TYPE ST_MotorData :
STRUCT
	bEnabled       : BOOL;                              // motor enabled
	fSpeedSetpoint : LREAL        := 0.0;
	nErrorCode     : UDINT;
	sName          : STRING(80)   := 'Motor';
	eState         : E_MotorState := E_MotorState.Idle; (* state *)
	counter        : INT;
END_STRUCT
END_TYPE

(* stored: Version 1.1.0.1
   DUT ST_MotorData: Id {bf3b27fe-277b-42e8-9d3c-5f37e955d5fb} *)
